TYPE "ST_FraktalHal"
VERSION : 0.1
   STRUCT
      "StationA" {ExternalAccessible := 'False'; ExternalVisible := 'False'; ExternalWritable := 'False'} : "ST_DeclarationUnitHal";
      "StationB" {ExternalAccessible := 'False'; ExternalVisible := 'False'; ExternalWritable := 'False'} : "ST_DeclarationUnitHal";
   END_STRUCT;
END_TYPE
